(* IEC 61131-3 sources: PLC-Static-Analysis/modules/plc-rules/src/test/resources/PLCA-P002, 2 files *)

(* ---- compliant.st ---- *)
PROGRAM P_IoOk
VAR
    iButton AT %IX0.0 : BOOL;
    qLamp AT %QX0.1 : BOOL;
    iTemp AT %I* : INT;
END_VAR
qLamp := iButton AND iTemp > 0;
END_PROGRAM

(* ---- noncompliant.st ---- *)
PROGRAM P_Io
VAR
    b : BOOL;
    w : WORD;
END_VAR
b := %IX0.0; // PLCA-P002
%QX0.1 := b; // PLCA-P002
w := %MW10 + %IW2; // PLCA-P002 PLCA-P002
END_PROGRAM
